// TIA Portal V21 export
VAR_GLOBAL   // PLC tag table "Default tag table"
   "Clock_2.5Hz" AT %M0.2 : Bool;
   Clock_5Hz AT %M0.1 : Bool;
   DiagStatusUpdate AT %M1.1 : Bool;
   "Clock_1.25Hz" AT %M0.4 : Bool;
   "Clock_0.625Hz" AT %M0.6 : Bool;
   AlwaysFALSE AT %M1.3 : Bool;
   FirstScan AT %M1.0 : Bool;
   "Clock_0.5Hz" AT %M0.7 : Bool;
   AlwaysTRUE AT %M1.2 : Bool;
   Clock_2Hz AT %M0.3 : Bool;
   Clock_Byte AT %MB0 : Byte;
   Clock_1Hz AT %M0.5 : Bool;
   System_Byte AT %MB1 : Byte;
   Clock_10Hz AT %M0.0 : Bool;
   ___testbool___ AT %M2.0 : Bool;
END_VAR
